{attribute 'Tc2GvlVarNames'}
VAR_GLOBAL CONSTANT
	nALARM_MAX_NO			:INT := 31;			(* Maximal number of alarms *)
END_VAR

(* stored: Version 1.1.0.1, ProductVersion 3.1.4024.15
   GVL GVL_FB_Alarm: Id {fc28ad4c-6b10-4499-aabe-93d931f52f89} *)
